# EPICS substitutions: db/Beckhoff_5XXX/ecmcEL5042.substitutions
file "ecmcEL5042-chX.template"
{
  pattern {CH_ID}
          {01   }
          {02   }
}
